Fanuc KAREL source: KA00077.KL

PROGRAM KA00077
%NOLOCKGROUP
VAR
  SRC: XYZWPREXT
  DST: POSITION
BEGIN
  SRC.X = 1.0
  DST = SRC
END KA00077
